(* IEC 61131-3 sources: Benedict-Informatik/Modul 319 Elektrotechnik/Leeres_Grundgeruest_mit_TON, 1 file *)

(* ---- Leeres_Grundgeruest_mit_TON_PLC_PRG.st ---- *)
PROGRAM PLC_PRG
VAR
	E1 : BOOL;
	E3 : BOOL;
	T1 : TON;
	K1 : BOOL;
END_VAR

(* Noch keine Logik implementiert *)
